(* IEC 61131-3 sources: RootPLC/conformance/cases/pous, 52 files *)

(* ---- err_missing_end.st ---- *)
(* spec: [pous.end]
   expect: error RP0202 *)
TYPE ST_Point :
STRUCT
    x : INT;
    y : INT;
END_STRUCT;

(* ---- ok_type_spec.st ---- *)
(* spec: [pous.type-block] [pous.type-spec]
   expect: ok *)
TYPE
    Percent : INT (0..100);
    Mode : (Off, Manual, Auto);
    Code : INT (Good := 0, Fail := 1);
    Name : STRING[20];
    Grid : ARRAY[1..3, 1..3] OF REAL;
    PInt : REF_TO INT;
    Pair : STRUCT
        a : INT;
        b : BOOL;
    END_STRUCT;
END_TYPE

(* ---- warn_interface_syntax.st ---- *)
(* spec: [pous.oop.interface] [scope.vendor-forms]
   expect: warning RP0134 *)
INTERFACE I_Base
METHOD Reset
END_METHOD
END_INTERFACE

INTERFACE I_Motor EXTENDS I_Base
METHOD Start : BOOL
VAR_INPUT
    speed : INT;
END_VAR
END_METHOD
PROPERTY Running : BOOL
END_PROPERTY
END_INTERFACE

(* ---- err_extends_not_fb.st ---- *)
(* spec: [pous.oop.extends]
   expect: error RP0111 *)
TYPE S : STRUCT a : INT; END_STRUCT; END_TYPE

FUNCTION_BLOCK FB_X EXTENDS S
END_FUNCTION_BLOCK

(* ---- err_fb_local_write.st ---- *)
(* spec: [pous.call.local-read]
   expect: error RP0203 *)
FUNCTION_BLOCK FB_Plant
VAR
    n : INT;
    arr : ARRAY[0..3] OF INT;
END_VAR
END_FUNCTION_BLOCK

PROGRAM PRG_Main
VAR
    fbPlant : FB_Plant;
END_VAR
fbPlant.n := 1;        (* internal variables are read-only from outside *)
fbPlant.arr[1] := 2;
END_PROGRAM

(* ---- err_interface_assign.st ---- *)
(* spec: [pous.oop.interface-ref]
   expect: error RP0103 *)
INTERFACE I_A
METHOD M : INT
END_METHOD
END_INTERFACE

FUNCTION_BLOCK FB_Z
END_FUNCTION_BLOCK

PROGRAM PRG_Main
VAR
    a : I_A;
    z : FB_Z;
END_VAR
a := z;
END_PROGRAM

(* ---- err_interface_not_implemented.st ---- *)
(* spec: [pous.oop.implements]
   expect: error RP0203 *)
INTERFACE I_A
METHOD M : INT
END_METHOD
END_INTERFACE

FUNCTION_BLOCK FB_X IMPLEMENTS I_A
END_FUNCTION_BLOCK

(* ---- err_no_result_in_expression.st ---- *)
(* spec: [pous.oop.method] [pous.function]
   expect: error RP0303 *)
(* A method without a result type has no value (found in a corpus block
   that assigned such a call; vendor compilers reject it). *)
FUNCTION_BLOCK FB_Buffer
VAR size : UDINT := 100; END_VAR
METHOD SetSize
VAR_INPUT n : UDINT; END_VAR
size := n;
END_METHOD
END_FUNCTION_BLOCK

PROGRAM PRG_Main
VAR
    b : FB_Buffer;
    n : UDINT := 32;
END_VAR
b.SetSize(n);
n := b.SetSize(n);
END_PROGRAM

(* ---- err_oop_downcast.st ---- *)
(* spec: [pous.oop.upcast]
   expect: error RP0103 *)
FUNCTION_BLOCK Product
END_FUNCTION_BLOCK

FUNCTION_BLOCK Chips EXTENDS Product
END_FUNCTION_BLOCK

PROGRAM PRG_Main
VAR
    b : Product;
    rb : REF_TO Product;
    rc : REF_TO Chips;
END_VAR
rb := REF(b);
rc := rb;
END_PROGRAM

(* ---- in_out_writes_back.st ---- *)
(* spec: [pous.call.in-out]
   expect: ok
   run: PRG_Main cycles=2
   assert: total = 10
   assert: count = 2
   assert: arr[2] = 4 *)
FUNCTION AddTo : BOOL
VAR_IN_OUT
    acc : INT;
END_VAR
VAR_INPUT
    n : INT;
END_VAR
acc := acc + n;
AddTo := TRUE;
END_FUNCTION

FUNCTION_BLOCK FB_Count
VAR_IN_OUT
    c : INT;
END_VAR
c := c + 1;
END_FUNCTION_BLOCK

PROGRAM PRG_Main
VAR
    total, count : INT;
    arr : ARRAY[1..3] OF INT;
    ok : BOOL;
    fb : FB_Count;
END_VAR
ok := AddTo(acc := total, n := 5);
fb(c := count);
ok := AddTo(arr[2], 2);
END_PROGRAM

(* ---- ok_action.st ---- *)
(* spec: [pous.action]
   expect: ok
   run: PRG_Main cycles=1
   assert: n = 3
   assert: m = 10 *)
FUNCTION_BLOCK FB_Counter
VAR_OUTPUT
    count : INT;
END_VAR
ACTION Reset:
    count := 0;
END_ACTION
ACTION Advance:
    count := count + 1;
END_ACTION
END_FUNCTION_BLOCK

FUNCTION_BLOCK FB_Tank
VAR_OUTPUT
    level : INT;
END_VAR
END_FUNCTION_BLOCK

ACTION Fill:
    level := 10;
END_ACTION

PROGRAM PRG_Main
VAR
    c : FB_Counter;
    t : FB_Tank;
    n, m : INT;
END_VAR
c.Advance();
c.Advance();
c.Reset();
c.Advance();
c.Advance();
c.Advance();
n := c.count;
t.Fill();
m := t.level;
END_PROGRAM

(* ---- ok_class.st ---- *)
(* spec: [pous.oop.class]
   expect: ok
   run: PRG_Main cycles=1
   assert: v = 6 *)
CLASS Accumulator
VAR
    sum : INT;
END_VAR
METHOD PUBLIC Add : INT
VAR_INPUT
    x : INT;
END_VAR
sum := sum + x;
Add := sum;
END_METHOD
END_CLASS

PROGRAM PRG_Main
VAR
    acc : Accumulator;
    v : INT;
END_VAR
acc.Add(x := 1);
acc.Add(x := 2);
v := acc.Add(x := 3);
END_PROGRAM

(* ---- ok_extends.st ---- *)
(* spec: [pous.oop.extends]
   expect: ok
   run: PRG_Main cycles=2
   assert: base_count = 2
   assert: own_count = 2 *)
FUNCTION_BLOCK FB_Counter
VAR_OUTPUT
    count : INT;
END_VAR
count := count + 1;
END_FUNCTION_BLOCK

FUNCTION_BLOCK FB_Pair EXTENDS FB_Counter
VAR_OUTPUT
    mine : INT;
END_VAR
SUPER^();
mine := mine + 1;
END_FUNCTION_BLOCK

PROGRAM PRG_Main
VAR
    p : FB_Pair;
    base_count, own_count : INT;
END_VAR
p();
base_count := p.count;
own_count := p.mine;
END_PROGRAM

(* ---- ok_function_block.st ---- *)
(* spec: [pous.function] [pous.function-block] [statements.call] [statements.assignment]
   expect: ok
   run: PRG_Main cycles=1
   assert: n = 1
   assert: y = 10 *)
FUNCTION Clamp : INT
VAR_INPUT
    v, lo, hi : INT;
END_VAR
IF v < lo THEN
    Clamp := lo;
ELSIF v > hi THEN
    Clamp := hi;
ELSE
    Clamp := v;
END_IF;
END_FUNCTION

FUNCTION_BLOCK FB_Counter
VAR_INPUT
    pulse : BOOL;
END_VAR
VAR_OUTPUT
    count : INT;
END_VAR
IF pulse THEN
    count := count + 1;
END_IF;
END_FUNCTION_BLOCK

PROGRAM PRG_Main
VAR
    c : FB_Counter;
    n : INT;
    y : INT;
END_VAR
c(pulse := TRUE, count => n);
y := Clamp(15, 0, 10);
END_PROGRAM

(* ---- ok_implements_syntax.st ---- *)
(* spec: [pous.oop.implements]
   expect: ok *)
INTERFACE I_Resettable
METHOD Reset
END_METHOD
END_INTERFACE

FUNCTION_BLOCK FB_Timer IMPLEMENTS I_Resettable
VAR
    t : INT;
END_VAR
METHOD Reset
t := 0;
END_METHOD
END_FUNCTION_BLOCK

(* ---- ok_in_out_same_variable.st ---- *)
(* spec: [pous.call.in-out]
   expect: ok
   run: PRG_Main cycles=1
   assert: viaFb = 2
   assert: viaFun = 3
   assert: seen = 3
   assert: shown = 2 *)
(* The counter keeps a pointer into itself; passed as VAR_IN_OUT, the
   write through that pointer and the parameter are one variable. *)
FUNCTION_BLOCK Counter
VAR_OUTPUT
    v : INT;
END_VAR
VAR
    p : REF_TO INT;
END_VAR
IF p = NULL THEN
    p := REF(v);
END_IF;
p^ := p^ + 1;
END_FUNCTION_BLOCK

FUNCTION_BLOCK Bump
VAR_IN_OUT
    c : Counter;
END_VAR
VAR_OUTPUT
    seen : INT;
END_VAR
c();
seen := c.v;
END_FUNCTION_BLOCK

FUNCTION BumpF : INT
VAR_IN_OUT
    c : Counter;
END_VAR
c();
BumpF := c.v;
END_FUNCTION

PROGRAM PRG_Main
VAR
    cnt : Counter;
    b : Bump;
    viaFb, viaFun, seen, shown : INT;
END_VAR
cnt();
b(c := cnt);
viaFb := cnt.v;
shown := b.seen;
seen := BumpF(cnt);
viaFun := cnt.v;
END_PROGRAM

(* ---- ok_in_out_through_action.st ---- *)
(* spec: [pous.call.in-out]
   expect: ok
   run: PRG_Main cycles=1
   assert: first = 1
   assert: second = 2
   assert: seen = 2 *)
TYPE ST_Steps :
STRUCT
    list : ARRAY[0..3] OF INT;
END_STRUCT;
END_TYPE

(* the action writes the block's VAR_IN_OUT: the caller's variable *)
FUNCTION_BLOCK StepFb
VAR_INPUT
    k : INT;
END_VAR
VAR_IN_OUT
    st : ST_Steps;
END_VAR
VAR_OUTPUT
    seen : INT;
END_VAR
Register();
seen := st.list[2];

ACTION Register:
st.list[k] := k;
END_ACTION
END_FUNCTION_BLOCK

FUNCTION_BLOCK Chain
VAR_IN_OUT
    st : ST_Steps;
END_VAR
VAR
    a, b : StepFb;
END_VAR
VAR_OUTPUT
    seen : INT;
END_VAR
a(k := 1, st := st);
b(k := 2, st := st);
seen := a.seen;
END_FUNCTION_BLOCK

PROGRAM PRG_Main
VAR
    c : Chain;
    s : ST_Steps;
    first, second, seen : INT;
END_VAR
c(st := s);
c(st := s);
first := s.list[1];
second := s.list[2];
seen := c.seen;
END_PROGRAM

(* ---- ok_interface_dispatch.st ---- *)
(* spec: [pous.oop.interface-ref]
   expect: ok
   run: PRG_Main cycles=1
   assert: total = 14
   assert: empty
   assert: set *)
INTERFACE I_Shape
METHOD Area : INT
END_METHOD
END_INTERFACE

FUNCTION_BLOCK FB_Square IMPLEMENTS I_Shape
VAR_INPUT
    side : INT := 2;
END_VAR
METHOD Area : INT
Area := side * side;
END_METHOD
END_FUNCTION_BLOCK

FUNCTION_BLOCK FB_Rect IMPLEMENTS I_Shape
VAR_INPUT
    w : INT := 2;
    h : INT := 5;
END_VAR
METHOD Area : INT
Area := w * h;
END_METHOD
END_FUNCTION_BLOCK

PROGRAM PRG_Main
VAR
    sq : FB_Square;
    re : FB_Rect;
    shapes : ARRAY[1..2] OF I_Shape;
    none : I_Shape;
    i, total : INT;
    empty, set : BOOL;
END_VAR
shapes[1] := sq;
shapes[2] := re;
FOR i := 1 TO 2 DO
    total := total + shapes[i].Area();
END_FOR;
empty := none = NULL;
set := shapes[1] <> NULL;
END_PROGRAM

(* ---- ok_methods.st ---- *)
(* spec: [pous.oop.method]
   expect: ok
   run: PRG_Main cycles=1
   assert: total = 7
   assert: r = 14 *)
FUNCTION_BLOCK FB_Acc
VAR
    sum : INT;
END_VAR
METHOD Add : INT
VAR_INPUT
    amount : INT;
END_VAR
sum := sum + amount;
Add := sum;
END_METHOD
METHOD Double : INT
Double := Add(amount := sum);
END_METHOD
END_FUNCTION_BLOCK

PROGRAM PRG_Main
VAR
    acc : FB_Acc;
    total, r : INT;
END_VAR
acc.Add(amount := 3);
total := acc.Add(amount := 4);
r := acc.Double();
END_PROGRAM

(* ---- ok_oop_modifiers.st ---- *)
(* spec: [pous.oop.modifiers]
   expect: ok
   run: PRG_Main cycles=1
   assert: v = 2 *)
FUNCTION_BLOCK PUBLIC FINAL FB_Two
METHOD PUBLIC Value : INT
Value := 2;
END_METHOD
METHOD PRIVATE Helper
END_METHOD
END_FUNCTION_BLOCK

PROGRAM PRG_Main
VAR
    t : FB_Two;
    v : INT;
END_VAR
v := t.Value();
END_PROGRAM

(* ---- ok_override_dispatch.st ---- *)
(* spec: [pous.oop.override]
   expect: ok
   run: PRG_Main cycles=1
   assert: a = 9
   assert: b = 9
   assert: c = 0 *)
FUNCTION_BLOCK FB_Shape
METHOD Area : INT
Area := 0;
END_METHOD
METHOD Describe : INT
Describe := Area();
END_METHOD
END_FUNCTION_BLOCK

FUNCTION_BLOCK FB_Square EXTENDS FB_Shape
VAR
    side : INT := 3;
END_VAR
METHOD OVERRIDE Area : INT
Area := side * side;
END_METHOD
METHOD Base : INT
Base := SUPER^.Area();
END_METHOD
END_FUNCTION_BLOCK

PROGRAM PRG_Main
VAR
    sq : FB_Square;
    a, b, c : INT;
END_VAR
a := sq.Area();
b := sq.Describe();
c := sq.Base();
END_PROGRAM

(* ---- ok_qualified_type.st ---- *)
(* spec: [pous.type-spec]
   expect: ok
   run: PRG_Main cycles=1
   assert: n = 3 *)
TYPE T_Count : INT; END_TYPE

FUNCTION_BLOCK FB_Base
VAR_OUTPUT
    n : MyLib.T_Count := 3;
END_VAR
END_FUNCTION_BLOCK

FUNCTION_BLOCK FB_Derived EXTENDS MyLib.FB_Base
END_FUNCTION_BLOCK

PROGRAM PRG_Main
VAR
    d : FB_Derived;
    n : INT;
END_VAR
n := d.n;
END_PROGRAM

(* ---- ok_test_block.st ---- *)
(* spec: [pous.test]
   expect: ok *)
FUNCTION_BLOCK FB_Latch
VAR_INPUT
    set, reset : BOOL;
END_VAR
VAR_OUTPUT
    q : BOOL;
END_VAR
q := (set OR q) AND NOT reset;
END_FUNCTION_BLOCK

TEST latch_sets
VAR
    uut : FB_Latch;
END_VAR
uut(set := TRUE);
ASSERT_TRUE(uut.q);
END_TEST

(* ---- ok_this_super.st ---- *)
(* spec: [pous.oop.this]
   expect: ok
   run: PRG_Main cycles=1
   assert: v = 5 *)
FUNCTION_BLOCK FB_Box
VAR
    hidden : INT;
END_VAR
METHOD Set
VAR_INPUT
    x : INT;
END_VAR
THIS^.hidden := x;
END_METHOD
METHOD Get : INT
Get := THIS^.hidden;
END_METHOD
END_FUNCTION_BLOCK

PROGRAM PRG_Main
VAR
    b : FB_Box;
    v : INT;
END_VAR
b.Set(x := 5);
v := b.Get();
END_PROGRAM

(* ---- warn_fb_init_local.st ---- *)
(* spec: [variables.init-arguments] [pous.oop.fb-init]
   expect: warning RP0119 RP0135 RP0134
   run: P cycles=2
   assert: s = 'made'
   assert: calls = 2 *)
VAR_GLOBAL
    inits : INT;
END_VAR

FUNCTION_BLOCK FB_Named
VAR_OUTPUT
    name : STRING;
END_VAR
METHOD FB_init : BOOL
VAR_INPUT
    bInitRetains : BOOL;
    bInCopyCode : BOOL;
    sName : STRING;
END_VAR
name := sName;
inits := inits + 1;
END_METHOD
END_FUNCTION_BLOCK

FUNCTION F_Make : STRING
VAR
    n : FB_Named('made');
END_VAR
F_Make := n.name;
END_FUNCTION

PROGRAM P
VAR
    s : STRING;
    calls : INT;
END_VAR
s := F_Make();
calls := inits;
END_PROGRAM

(* ---- warn_fb_init_registry.st ---- *)
(* spec: [pous.oop.fb-init] [pous.oop.override] [scope.vendor-forms]
   expect: warning RP0135 RP0116 RP0134
   run: PRG_Main cycles=2
   assert: a.hits = 2
   assert: b.hits = 4
   assert: seen = 12 *)
VAR_GLOBAL
    count : UINT;
    order : INT;
    suites : ARRAY[1..4] OF POINTER TO FB_Suite;
END_VAR

(* a TcUnit-style registry: every instance registers itself in FB_init,
   and a runner calls each body through a pointer of the base type *)
FUNCTION_BLOCK FB_Suite
VAR
    hits : INT;
    id : INT;
END_VAR
METHOD FB_init : BOOL
VAR_INPUT
    bInitRetains : BOOL;
    bInCopyCode : BOOL;
END_VAR
count := count + 1;
id := UINT_TO_INT(count);
order := order * 10 + id;
suites[count] := THIS;
END_METHOD
METHOD Tick
hits := hits + 1;
END_METHOD
END_FUNCTION_BLOCK

FUNCTION_BLOCK FB_Single EXTENDS FB_Suite
Tick();
END_FUNCTION_BLOCK

FUNCTION_BLOCK FB_Double EXTENDS FB_Suite
METHOD Tick
hits := hits + 2;
END_METHOD
Tick();
END_FUNCTION_BLOCK

PROGRAM PRG_Main
VAR
    b : FB_Double;
    a : FB_Single;
    i : UINT;
    seen : INT;
END_VAR
seen := order;
FOR i := 1 TO count DO
    suites[i]^();
END_FOR;
END_PROGRAM

(* ---- warn_fb_local_read.st ---- *)
(* spec: [pous.call.local-read]
   expect: warning RP0130
   run: PRG_Main cycles=1
   assert: a = 3
   assert: b = 4
   assert: c = 30
   assert: d = 7 *)
FUNCTION_BLOCK FB_Inner
VAR
    nCount : INT := 3;
END_VAR
METHOD Bump : INT
nCount := nCount + 1;
Bump := nCount;
END_METHOD
END_FUNCTION_BLOCK

FUNCTION_BLOCK FB_Plant
VAR
    fbInner : FB_Inner;
    arr : ARRAY[0..3] OF INT := [10, 20, 30, 40];
END_VAR
END_FUNCTION_BLOCK

PROGRAM PRG_Main
VAR
    fbPlant : FB_Plant;
    a, b, c, d : INT;
    out : ARRAY[0..5] OF INT;
END_VAR
a := fbPlant.fbInner.nCount;        (* read an internal variable *)
b := fbPlant.fbInner.Bump();        (* call a method of an internal instance *)
c := fbPlant.arr[2];                (* read an element of an internal array *)
out[fbPlant.fbInner.nCount] := 7;   (* a read inside an assignment target *)
d := out[4];
END_PROGRAM

(* ---- warn_header_semicolon.st ---- *)
(* spec: [pous.function-block] [scope.vendor-forms]
   expect: warning RP0134
   run: PRG_Main cycles=1
   assert: v = 7 *)
FUNCTION Seven : INT;
Seven := 7;
END_FUNCTION

FUNCTION_BLOCK FB_X
METHOD Get : INT;
VAR_INPUT
    x : INT;
END_VAR
Get := x;
END_METHOD
END_FUNCTION_BLOCK

PROGRAM PRG_Main
VAR
    f : FB_X;
    v : INT;
END_VAR
v := f.Get(x := Seven());
END_PROGRAM

(* ---- warn_interface_zero_init.st ---- *)
(* spec: [pous.oop.interface-ref] [scope.vendor-forms]
   expect: warning RP0127
   run: PRG_Main cycles=1
   assert: a = TRUE
   assert: b = TRUE
   assert: c = 5 *)
INTERFACE I_Value
METHOD Get : INT
END_METHOD
END_INTERFACE

FUNCTION_BLOCK FB_Five IMPLEMENTS I_Value
METHOD Get : INT
Get := 5;
END_METHOD
END_FUNCTION_BLOCK

FUNCTION F_Read : INT
VAR_INPUT
    ip : I_Value := 0;
END_VAR
IF ip <> 0 THEN
    F_Read := ip.Get();
END_IF;
END_FUNCTION

PROGRAM PRG_Main
VAR
    ipA : I_Value := 0;
    ipB : I_Value := NULL;
    five : FB_Five;
    a, b : BOOL;
    c : INT;
END_VAR
a := ipA = 0;
b := ipB = NULL AND F_Read() = 0;
c := F_Read(five);
END_PROGRAM

(* ---- warn_oop_accessor_modifiers.st ---- *)
(* spec: [pous.oop.modifiers] [scope.vendor-forms]
   expect: warning RP0134
   run: PRG_Main cycles=1
   assert: x = 9 *)
FUNCTION_BLOCK FB_Store
VAR
    v : INT := 4;
END_VAR
PROPERTY PUBLIC Value : INT
GET PUBLIC
    Value := v;
END_GET
SET PROTECTED
    v := Value;
END_SET
END_PROPERTY
END_FUNCTION_BLOCK

PROGRAM PRG_Main
VAR
    f : FB_Store;
    x : INT;
END_VAR
f.Value := 9;
x := f.Value;
END_PROGRAM

(* ---- warn_oop_upcast.st ---- *)
(* spec: [pous.oop.upcast] [types.reference.alias]
   expect: warning RP0118
   run: PRG_Main cycles=1
   assert: viaRef = 2
   assert: viaParam = 2
   assert: viaBase = 1
   assert: count = 2 *)
FUNCTION_BLOCK Product
VAR_OUTPUT
    taken : INT;
END_VAR
METHOD Price : INT
Price := 1;
END_METHOD
METHOD Take
taken := taken + 1;
END_METHOD
END_FUNCTION_BLOCK

FUNCTION_BLOCK Chips EXTENDS Product
METHOD Price : INT
Price := 2;
END_METHOD
END_FUNCTION_BLOCK

FUNCTION_BLOCK Snack EXTENDS Chips
END_FUNCTION_BLOCK

FUNCTION PriceOf : INT
VAR_INPUT
    p : REFERENCE TO Product;
END_VAR
p.Take();
PriceOf := p.Price();
END_FUNCTION

PROGRAM PRG_Main
VAR
    s : Snack;
    b : Product;
    r : REF_TO Product;
    viaRef, viaParam, viaBase, count : INT;
END_VAR
r := REF(s);
viaRef := r^.Price();
viaParam := PriceOf(s);
viaBase := PriceOf(b);
r^.Take();
count := s.taken;
END_PROGRAM

(* ---- warn_property_access.st ---- *)
(* spec: [pous.oop.property] [scope.vendor-forms]
   expect: warning RP0134
   run: PRG_Main cycles=1
   assert: a = 40
   assert: b = 50
   assert: c = 7
   assert: d = 14 *)
INTERFACE I_Level
PROPERTY Level : INT
GET
END_GET
END_PROPERTY
END_INTERFACE

FUNCTION_BLOCK FB_Valve IMPLEMENTS I_Level
VAR
    pos : INT;
END_VAR
PROPERTY Position : INT
GET
    Position := pos;
END_GET
SET
    pos := LIMIT(0, Position, 100);
END_SET
END_PROPERTY
PROPERTY Level : INT
GET
    Level := pos;
END_GET
END_PROPERTY
METHOD Open
Position := Position + 10;
END_METHOD
END_FUNCTION_BLOCK

FUNCTION_BLOCK FB_Doubler EXTENDS FB_Valve
PROPERTY Level : INT
GET
    Level := SUPER^.Level * 2;
END_GET
END_PROPERTY
END_FUNCTION_BLOCK

PROGRAM PRG_Main
VAR
    v : FB_Valve;
    w : FB_Doubler;
    itf : I_Level;
    a, b, c, d : INT;
END_VAR
v.Position := 30;
v.Open();
a := v.Position;
v.Position := v.Position + 10;
b := v.Level;
w.Position := 7;
itf := w;
c := w.Position;
d := itf.Level;
END_PROGRAM

(* ---- warn_property_named_set.st ---- *)
(* spec: [pous.oop.property] [scope.vendor-forms]
   expect: warning RP0134
   run: PRG_Main cycles=1
   assert: v = 2.5 *)
FUNCTION_BLOCK FB_Control
VAR
    fSet : REAL;
END_VAR
PROPERTY Set : REAL
GET
    Set := fSet;
END_GET
SET
    fSet := Set;
END_SET
END_PROPERTY
END_FUNCTION_BLOCK

PROGRAM PRG_Main
VAR
    c : FB_Control;
    v : REAL;
END_VAR
c.Set := 2.5;
v := c.Set;
END_PROGRAM

(* ---- warn_property_syntax.st ---- *)
(* spec: [pous.oop.property] [scope.vendor-forms]
   expect: warning RP0134 *)
FUNCTION_BLOCK FB_Valve
VAR
    pos : INT;
END_VAR
PROPERTY Position : INT
GET
    Position := pos;
END_GET
SET
    pos := Position;
END_SET
END_PROPERTY
END_FUNCTION_BLOCK

(* ---- warn_var_inst.st ---- *)
(* spec: [pous.oop.method] [scope.vendor-forms]
   expect: warning RP0134
   run: PRG_Main cycles=3
   assert: a = 3
   assert: b = 3 *)
FUNCTION_BLOCK FB_Counter
METHOD Next : INT
VAR_INST
    calls : INT;
END_VAR
calls := calls + 1;
Next := calls;
END_METHOD
END_FUNCTION_BLOCK

PROGRAM PRG_Main
VAR
    c1, c2 : FB_Counter;
    a, b : INT;
END_VAR
a := c1.Next();
b := c2.Next();
END_PROGRAM

(* ---- err_call_not_callable.st ---- *)
(* spec: [pous.call.callee]
   expect: error RP0132 *)
PROGRAM PRG_Main
VAR
    b : BOOL;
    i : INT;
END_VAR
i := b(1);   (* b is a variable, not a function *)
END_PROGRAM

(* ---- err_in_out_constant.st ---- *)
(* spec: [pous.call.in-out]
   expect: error RP0114 *)
FUNCTION AddTo : BOOL
VAR_IN_OUT
    acc : INT;
END_VAR
acc := acc + 1;
AddTo := TRUE;
END_FUNCTION

PROGRAM PRG_Main
VAR
    ok : BOOL;
END_VAR
ok := AddTo(acc := 5);
END_PROGRAM

(* ---- err_syntax.st ---- *)
(* spec: [syntax.general]
   expect: error RP0201 *)
PROGRAM PRG_Main
VAR
    x : INT;
END_VAR
x := ;
END_PROGRAM

(* ---- err_two_errors.st ---- *)
(* spec: [syntax.recovery]
   expect: error RP0301 RP0201 *)
PROGRAM PRG_Main
VAR
    x, y : INT;
END_VAR
x := 1
y := * 2;
END_PROGRAM

(* ---- in_out_string_whole_text.st ---- *)
(* spec: [pous.call.in-out]
   expect: ok
   run: PRG_Main cycles=1
   assert: n = 120
   assert: m = 120
   assert: k = 12 *)
FUNCTION F_Append : INT
VAR_IN_OUT
    s : STRING;
END_VAR
F_Append := LEN(s);
s := CONCAT(s, 'abcdefghij');
END_FUNCTION

PROGRAM PRG_Main
VAR
    t : STRING[200];
    small : STRING[12] := 'xy';
    n, m, k : INT;
END_VAR
t := CONCAT('012345678901234567890123456789012345678901234567890123456789', '012345678901234567890123456789012345678901234567890123456789');
n := F_Append(t);
m := LEN(t) - 10;
F_Append(small);
k := LEN(small);
END_PROGRAM

(* ---- ok_call_function_shadowed_by_variable.st ---- *)
(* spec: [pous.call.callee]
   expect: ok
   run: PRG_Main cycles=1
   assert: r.Twice = 8 *)
FUNCTION Twice : INT
VAR_INPUT
    x : INT;
END_VAR
Twice := 2 * x;
END_FUNCTION

TYPE ST_R :
STRUCT
    Twice : INT;   (* a member named like the function *)
END_STRUCT;
END_TYPE

PROGRAM PRG_Main
VAR
    r : ST_R;
    Twice : STRING;   (* a variable named like the function *)
END_VAR
r.Twice := Twice(4);   (* calls the function *)
END_PROGRAM

(* ---- ok_function_body_at_once.st ---- *)
(* spec: [pous.function] [scope.vendor-forms]
   expect: warning RP0113 RP0134
   run: PRG_Main cycles=1
   assert: n = 2 *)
VAR_GLOBAL
    total : INT;
END_VAR

FUNCTION Bump
total := total + 1;
END_FUNCTION

PROGRAM PRG_Main
VAR
    n : INT;
END_VAR
Bump();
Bump();
n := total;
END_PROGRAM

(* ---- ok_in_out_address.st ---- *)
(* spec: [pous.call.in-out]
   expect: ok
   run: PRG_Main cycles=1
   assert: seen = 42
   assert: value = 43 *)
FUNCTION AddressOf : REF_TO INT
VAR_IN_OUT
    x : INT;
END_VAR
AddressOf := REF(x);
END_FUNCTION

PROGRAM PRG_Main
VAR
    value : INT := 42;
    p : REF_TO INT;
    seen : INT;
END_VAR
p := AddressOf(value);
seen := p^;
p^ := 43;
END_PROGRAM

(* ---- ok_namespace.st ---- *)
(* spec: [pous.namespace]
   expect: ok
   run: PRG_Main cycles=1
   assert: v = 4 *)
NAMESPACE Plant.Utils
FUNCTION Twice : INT
VAR_INPUT
    x : INT;
END_VAR
Twice := 2 * x;
END_FUNCTION
END_NAMESPACE

USING Plant.Utils;

PROGRAM PRG_Main
VAR
    v : INT;
END_VAR
v := Twice(x := 2);
END_PROGRAM

(* ---- ok_test_as_name.st ---- *)
(* spec: [pous.test]
   expect: ok
   run: PRG_Main cycles=1
   assert: n = 2 *)
FUNCTION TEST : INT
VAR_INPUT
    name : STRING;
END_VAR
TEST := LEN(name);
END_FUNCTION

PROGRAM PRG_Main
VAR
    n : INT;
END_VAR
n := TEST('ab');
END_PROGRAM

(* ---- ok_test_variable.st ---- *)
(* spec: [pous.test]
   expect: ok
   run: PRG_Main cycles=1
   assert: n = 4 *)
FUNCTION Twice : INT
VAR_INPUT
    x : INT;
END_VAR
VAR
    Test : INT;
END_VAR
Test := 2 * x;
Twice := Test;
END_FUNCTION

PROGRAM PRG_Main
VAR
    n : INT;
END_VAR
n := Twice(x := 2);
END_PROGRAM

(* ---- warn_function_modifier.st ---- *)
(* spec: [pous.oop.modifiers]
   expect: warning RP0124
   run: PRG_Main cycles=1
   assert: a = 6
   assert: b = 4.0 *)
FUNCTION INTERNAL F_Triple : INT
VAR_INPUT
    x : INT;
END_VAR
F_Triple := x * 3;
END_FUNCTION

FUNCTION OVERRIDE : REAL
VAR_INPUT
    x : REAL;
END_VAR
OVERRIDE := x * 2.0;
END_FUNCTION

PROGRAM PRG_Main
VAR
    a : INT;
    b : REAL;
END_VAR
a := F_Triple(2);
b := OVERRIDE(2.0);
END_PROGRAM

(* ---- warn_function_without_result.st ---- *)
(* spec: [pous.function]
   expect: warning RP0113
   run: PRG_Main cycles=2
   assert: total = 10 *)
FUNCTION AddTo
VAR_IN_OUT
    acc : INT;
END_VAR
VAR_INPUT
    n : INT;
END_VAR
acc := acc + n;
END_FUNCTION

PROGRAM PRG_Main
VAR
    total : INT;
END_VAR
AddTo(acc := total, n := 5);
END_PROGRAM

(* ---- warn_in_out_constant_value.st ---- *)
(* spec: [pous.call.in-out-constant] [scope.vendor-forms]
   expect: warning RP0134
   run: PRG_Main cycles=1
   assert: a = 3
   assert: b = 4
   assert: c = 9 *)
FUNCTION F_Len : INT
VAR_IN_OUT CONSTANT
    s : STRING;
END_VAR
F_Len := LEN(s);
END_FUNCTION

PROGRAM PRG_Main
VAR
    a, b, c : INT;
    t : STRING := 'abcd';
END_VAR
a := F_Len('xyz');
b := F_Len(t);
c := F_Len(CONCAT(t, 'efghi'));
END_PROGRAM

(* ---- warn_namespace_nested.st ---- *)
(* spec: [pous.namespace] [scope.vendor-forms]
   expect: warning RP0134
   run: PRG_Main cycles=1
   assert: a = 10
   assert: b = 10
   assert: ok = TRUE *)
NAMESPACE Lib
NAMESPACE Params
VAR_GLOBAL CONSTANT
    MaxSuites : UINT := 10;
END_VAR
END_NAMESPACE
FUNCTION Check : BOOL
VAR_INPUT n : UINT; END_VAR
Check := n > 0;
END_FUNCTION
END_NAMESPACE

PROGRAM PRG_Main
VAR
    a, b : UINT;
    ok : BOOL;
END_VAR
a := Lib.Params.MaxSuites;
b := Params.MaxSuites;
ok := Lib.Check(a);
END_PROGRAM

(* ---- warn_pou_closed_by_eof.st ---- *)
(* spec: [pous.end]
   expect: warning RP0131 *)
(* a CODESYS object export: the program has no END_PROGRAM; the end of
   the file closes it *)
PROGRAM PRG_Main
VAR
    n : INT;
END_VAR
n := n + 1;

(* ---- warn_stray_semicolons.st ---- *)
(* spec: [pous.stray-semicolon] [variables.declaration] [scope.vendor-forms]
   expect: warning RP0134
   run: PRG_Main cycles=1
   assert: x = 2
   assert: s.b = TRUE *)
TYPE E_Mode : (Idle, Run); END_TYPE;

TYPE ST_Pair :
STRUCT
    a : INT;;
    b : BOOL := TRUE;
END_STRUCT
END_TYPE

PROGRAM PRG_Main
VAR
    x : INT := 1;;
    m : E_Mode;
    s : ST_Pair;
END_VAR
x := x + 1;
END_PROGRAM;
